(* IEC 61131-3 sources: volt/packages/volt-lsp-iec/test-corpus/pro2193/Device/Plc Logic/Application/09 Misc/Library Manager/L_SUDP_SlaveUpDownloadManager, 64 files *)

(* ---- L_SEMP_ITF_EVENTPARAMETERS.dut ---- *)
TYPE L_SEMP_ITF_EVENTPARAMETERS :
STRUCT
	EVENTPARAMETERS : ARRAY [0..1] OF L_SEMP_ITF_ParameterItem;
END_STRUCT
END_TYPE

(* ---- L_SEMP_ITF_PARAMETERITEM.dut ---- *)
TYPE L_SEMP_ITF_PARAMETERITEM :
STRUCT
	SIZE : BYTE;
	ETYPE : INT;
	VALUE : L_SEMP_ITF_ParaValue;
END_STRUCT
END_TYPE

(* ---- L_SEMP_ITF_PARAVALUE.dut ---- *)
TYPE L_SEMP_ITF_PARAVALUE :
UNION
	DWVALUE : DWORD;
	DNVALUE : DINT;
	FVALUE : REAL;
	STVALUE : STRING;
	DWTEXTLISTID : DWORD;
END_UNION
END_TYPE

(* ---- L_SUDP_BUS_TYPE.dut ---- *)
TYPE L_SUDP_BUS_TYPE :
(
	BUS_CAN := 15,
	BUS_ETC := 64
);
END_TYPE

(* ---- L_SUDP_CONTROL.dut ---- *)
TYPE L_SUDP_CONTROL :
(
	NONE := 0,
	CHECKVERSION := 1,
	DOWNLOAD := 2,
	UPLOAD := 3,
	RESTARTDEVICE := 4,
	PROVIDENEWPARSETCHECKSUM := 5,
	ONLINEPARADOWNLOAD := 6,
	RESTARTDEVICE2 := 7,
	RESTARTDEVICEI750 := 8,
	ABORT := 10
);
END_TYPE

(* ---- L_SUDP_CPAR_FILE_HDR.dut ---- *)
TYPE L_SUDP_CPAR_FILE_HDR :
STRUCT
	DWFILETYPE : DWORD;
	DWVERSION : DWORD;
	DWFILESIZE : DWORD;
	DWVENDOR : DWORD;
	DWPRODUCTTYPE : DWORD;
	DWREVISION : DWORD;
	DWDATAOFF : DWORD;
	DWDATASIZE : DWORD;
	DWFILECRC : DWORD;
END_STRUCT
END_TYPE

(* ---- L_SUDP_ERRORCODES.dut ---- *)
TYPE L_SUDP_ERRORCODES :
(
	NO_ERROR := 0,
	FILE_NOT_FOUND := 1,
	FILE_READ_ERROR := 2,
	PARAM_WRITE_ERROR := 4,
	SLAVE_ERROR := 5,
	PARA_FILE_TYPE_INVALID := 7,
	PARAM_READ_ERROR := 8,
	NO_BUFFER := 9,
	NO_MEMORY := 10,
	WRONG_VERSION_FORMAT := 11,
	ETC_STATE_COULD_NOT_BE_CHANGED := 12,
	GET_FIRMWARE_BINARY_FILE_NAME_FAILED := 13,
	SLAVE_FIRMWARE_UPDATE_FAILED := 14,
	PARAM_SET_UPDATE_FAILED := 15,
	PARAM_SET_FILE_UPLOAD_FAILED := 16,
	PARAM_UPLOAD_FILE_CREATE_FAILED := 17,
	PARAM_WRITE_TO_FILE_FAILED := 18,
	NO_CONFIG_INFORMATION := 19,
	NO_CURRENT_IEC_TASK_INFORMATION := 20,
	NO_FREE_ASYNC_MANAGER := 21,
	FILE_WRITE_ERROR := 22,
	SLAVE_FIRMWARE_UPDATE_HW_INCOMPATIBILITY := 23,
	ERROR_PARAMETERST_UPDATE_FAILED_PARAM_WRITE_ERRORS := 24,
	PARAM_DL_ERROR_FILE_READ_ERROR := 25,
	SLAVE_FW_UPDATE_HW_DIFFERS_NOT_UPDATED := 26
);
END_TYPE

(* ---- L_SUDP_ERRORINDEXSUBINDEX.dut ---- *)
TYPE L_SUDP_ERRORINDEXSUBINDEX :
STRUCT
	WINDEX : WORD;
	WSUBINDEX : BYTE;
END_STRUCT
END_TYPE

(* ---- L_SUDP_MAX_STRING_LENGTH.dut ---- *)
TYPE L_SUDP_MAX_STRING_LENGTH :
(
	FILE_NAME := 50,
	DEVICE_FIRMWARE_VERSION_NUMBER := 30,
	PATH_AND_FILE_NAME := 250,
	FILE_PATH := 200
);
END_TYPE

(* ---- L_SUDP_PAR_DATA_HDR.dut ---- *)
TYPE L_SUDP_PAR_DATA_HDR :
STRUCT
	DWPARTYPE : DWORD;
	DWPARDATAOFF : DWORD;
	DWPARDATSIZE : DWORD;
END_STRUCT
END_TYPE

(* ---- L_SUDP_PAR_FILE_HDR.dut ---- *)
TYPE L_SUDP_PAR_FILE_HDR :
STRUCT
	DWFILETYPE : DWORD;
	DWVERSION : DWORD;
	DWFILESIZE : DWORD;
	DWVENDOR : DWORD;
	DWPRODUCTTYPE : DWORD;
	DWREVISION : DWORD;
	DWDATAOFF : DWORD;
	DWDATASIZE : DWORD;
	DWFILECRC : DWORD;
END_STRUCT
END_TYPE

(* ---- L_SUDP_PAR_FILE_HDR_SEL_PS.dut ---- *)
TYPE L_SUDP_PAR_FILE_HDR_SEL_PS :
STRUCT
	DWFILETYPE : DWORD;
	DWVERSION : DWORD;
	DWFILESIZE : DWORD;
	DWFILECRC : DWORD;
	DWCOUNTPARAMETERSETS : DWORD;
	APARAMETERSETINFO : ARRAY [0..10] OF L_SUDP_PAR_FILE_HDR_SEL_PS_INFO;
END_STRUCT
END_TYPE

(* ---- L_SUDP_PAR_FILE_HDR_SEL_PS_INFO.dut ---- *)
TYPE L_SUDP_PAR_FILE_HDR_SEL_PS_INFO :
STRUCT
	DWPARAMETERSETNUMBER : DWORD;
	DWDATAOFFSET : DWORD;
END_STRUCT
END_TYPE

(* ---- L_SUDP_PARM_ERROR_CODE.dut ---- *)
TYPE L_SUDP_PARM_ERROR_CODE :
STRUCT
	DWERRORCODE : DWORD;
	WINDEX : WORD;
	WSUBINDEX : WORD;
END_STRUCT
END_TYPE

(* ---- L_SUDP_PARM_HDR.dut ---- *)
TYPE L_SUDP_PARM_HDR :
STRUCT
	U16SIZE : UINT;
	U16INDEX : UINT;
	U16SUBINDEX : UINT;
END_STRUCT
END_TYPE

(* ---- L_SUDP_PARM_RECORD.dut ---- *)
TYPE L_SUDP_PARM_RECORD :
STRUCT
	U16SIZE : UINT;
	U16INDEX : UINT;
	U16SUBINDEX : UINT;
	U8DATA : BYTE;
END_STRUCT
END_TYPE

(* ---- L_SUDP_PRM_FILE_READWRITE_STATES.dut ---- *)
TYPE L_SUDP_PRM_FILE_READWRITE_STATES :
(
	NONE,
	WAIT_FILE_SIZE,
	WAIT_READ_FILE_OPEN,
	READ_FILE_HEADERS,
	WRITE_FILE_HEADERS,
	WAIT_WRITE_FILE_OPEN,
	WAIT_READ_PARAM_HEADER,
	WAIT_READ_PARAM_VALUE,
	WAIT_READ_NEXT_PARAM_HEADER_AND_PARAM_VALUE,
	WAIT_WRITE_FILE_PARAMETER,
	WAIT_SET_NEW_FILE_POS_FOR_WRITE_HEADERS,
	WAIT_WRITE_NEW_FILE_HEADERS,
	WAIT_CALC_CHECKSUM,
	WAIT_DELETE_OLD_FILE,
	WAIT_RENAME_NEW_TO_OLD_FILE,
	CLOSE_READ_FILE,
	CLOSE_WRITE_FILE,
	DONE,
	ERROR
);
END_TYPE

(* ---- L_SUDP_STATE.dut ---- *)
TYPE L_SUDP_STATE :
(
	NONE := 0,
	ISREGISTERED := 1,
	DOWNLOADISNECESSARY := 2,
	DOWNLOADISNOTNECESSARY := 3,
	ISBUSY := 4,
	UPDOWNLOADDONE := 5,
	RESTARTDONE := 6,
	NEWCHECKSUMPROVIDED := 7,
	RESTARTDONE2 := 8,
	RESTARTDONEI750 := 9,
	ERROR := 10,
	ABORTED := 20
);
END_TYPE

(* ---- L_SUDP_SUCCESSCODES.dut ---- *)
TYPE L_SUDP_SUCCESSCODES :
(
	SLAVE_FIRMWARE_UPDATE_DONE := 1000,
	SHOW_OLD_FIRMWARE_VERSION := 2000,
	SUDP_DEBUG := 16#2003,
	SUDP_SLAVE_NOT_PRESENT := 16#2004
);
END_TYPE

(* ---- L_SUDP_TRANSFERTYPE.dut ---- *)
TYPE L_SUDP_TRANSFERTYPE :
(
	PARAMETERSETDOWNLOAD := 0,
	PARAMETERSETUPLOAD := 1,
	FIRMWAREDOWNLOAD := 2,
	FIRMWAREDOWNLOAD2 := 3,
	FIRMWAREDOWNLOADI750 := 4
);
END_TYPE

(* ---- DECIMALTOHEXSTRING.pou ---- *)
FUNCTION DECIMALTOHEXSTRING : STRING
VAR_INPUT
	DWVALUE : DWORD;
	NMAXBYTESIZE : INT;
END_VAR
END_FUNCTION

(* ---- GETBOOLEANPROPERTY.pou ---- *)
FUNCTION GETBOOLEANPROPERTY : BOOL
VAR_INPUT
	STKEY : WSTRING;
END_VAR
END_FUNCTION

(* ---- GETCOMPANY.pou ---- *)
FUNCTION GETCOMPANY : WSTRING
END_FUNCTION

(* ---- GETNUMBERPROPERTY.pou ---- *)
FUNCTION GETNUMBERPROPERTY : DINT
VAR_INPUT
	STKEY : WSTRING;
END_VAR
END_FUNCTION

(* ---- GETTEXTPROPERTY.pou ---- *)
FUNCTION GETTEXTPROPERTY : WSTRING
VAR_INPUT
	STKEY : WSTRING;
END_VAR
END_FUNCTION

(* ---- GETTEXTPROPERTY2.pou ---- *)
FUNCTION GETTEXTPROPERTY2 : POINTER TO WSTRING
VAR_INPUT
	STKEY : WSTRING;
END_VAR
END_FUNCTION

(* ---- GETTITLE.pou ---- *)
FUNCTION GETTITLE : WSTRING
END_FUNCTION

(* ---- GETVERSION.pou ---- *)
FUNCTION GETVERSION : VERSION
END_FUNCTION

(* ---- GETVERSIONPROPERTY.pou ---- *)
FUNCTION GETVERSIONPROPERTY : VERSION
VAR_INPUT
	STKEY : WSTRING;
END_VAR
END_FUNCTION

(* ---- L_EXISTALLFILES.pou ---- *)
FUNCTION L_EXISTALLFILES : BOOL
END_FUNCTION

(* ---- L_PATHFIRMWAREFILES.pou ---- *)
FUNCTION L_PATHFIRMWAREFILES : STRING(L_SUDP_MAX_STRING_LENGTH.FILE_PATH)
END_FUNCTION

(* ---- L_PATHPARAMETERSETFILES.pou ---- *)
FUNCTION L_PATHPARAMETERSETFILES : STRING(L_SUDP_MAX_STRING_LENGTH.FILE_PATH)
END_FUNCTION

(* ---- L_SUDP_CRC32FINISH.pou ---- *)
FUNCTION L_SUDP_CRC32FINISH : DWORD
VAR_INPUT
	ULCRC : DWORD;
END_VAR
END_FUNCTION

(* ---- L_SUDP_CRC32INIT.pou ---- *)
FUNCTION L_SUDP_CRC32INIT : DWORD
END_FUNCTION

(* ---- L_SUDP_CRC32UPDATE.pou ---- *)
FUNCTION L_SUDP_CRC32UPDATE : DWORD
VAR_INPUT
	ULCRC : DWORD;
	PDATA : POINTER TO BYTE;
	ULSIZE : __XWORD;
END_VAR
END_FUNCTION

(* ---- L_SUDP_GETBINARYFILENAME.pou ---- *)
FUNCTION L_SUDP_GETBINARYFILENAME : BOOL
VAR_INPUT
	WFIELDBUSMASTERID : WORD;
	WINTERFACE : WORD;
	DNNODEADDRESS : DINT;
	PSBINARYFILENAME : POINTER TO STRING(20);
END_VAR
END_FUNCTION

(* ---- L_SUDP_GETBUFFERINDEX.pou ---- *)
FUNCTION L_SUDP_GETBUFFERINDEX : WORD
VAR_INPUT
	DWLENGTH : DWORD;
	DWTASKINTERVAL : DWORD;
	PERROR : POINTER TO L_SUDP_ErrorCodes;
END_VAR
END_FUNCTION

(* ---- L_SUDP_GETFBCONTROL.pou ---- *)
FUNCTION L_SUDP_GETFBCONTROL : L_SUDP_Control
VAR_INPUT
	HREGISTRATION : CAA.HANDLE;
END_VAR
END_FUNCTION

(* ---- L_SUDP_GETFWDLMODE.pou ---- *)
FUNCTION L_SUDP_GETFWDLMODE : BYTE
END_FUNCTION

(* ---- L_SUDP_GETLEMREGISTRATIONHANDLE.pou ---- *)
FUNCTION L_SUDP_GETLEMREGISTRATIONHANDLE : RTS_IEC_HANDLE
END_FUNCTION

(* ---- L_SUDP_GETPATHBOOTDIRECTORY.pou ---- *)
FUNCTION L_SUDP_GETPATHBOOTDIRECTORY : STRING(L_SUDP_MAX_STRING_LENGTH.FILE_PATH)
END_FUNCTION

(* ---- L_SUDP_GETPATHTEMPDIRECTORY.pou ---- *)
FUNCTION L_SUDP_GETPATHTEMPDIRECTORY : STRING(L_SUDP_MAX_STRING_LENGTH.FILE_PATH)
END_FUNCTION

(* ---- L_SUDP_GETPOINTERTOBUFFER.pou ---- *)
FUNCTION L_SUDP_GETPOINTERTOBUFFER : POINTER TO BYTE
VAR_INPUT
	WBUFFERNUMBER : WORD;
	PERROR : POINTER TO L_SUDP_ErrorCodes;
END_VAR
END_FUNCTION

(* ---- L_SUDP_GETTARGETVERSION.pou ---- *)
FUNCTION L_SUDP_GETTARGETVERSION : BOOL
VAR_INPUT
	ETRANSFERTYPE : L_SUDP_TransferType;
	WFIELDBUSMASTERID : WORD;
	WINTERFACE : WORD;
	DNNODEADDRESS : DINT;
	PSTARGETVERSION : POINTER TO STRING(20);
END_VAR
END_FUNCTION

(* ---- L_SUDP_ISBOOTAPPLICATIONLOADED.pou ---- *)
FUNCTION L_SUDP_ISBOOTAPPLICATIONLOADED : BOOL
END_FUNCTION

(* ---- L_SUDP_REGISTER.pou ---- *)
FUNCTION L_SUDP_REGISTER : CAA.HANDLE
VAR_INPUT
	ETRANSFERTYPE : L_SUDP_TransferType;
	WFIELDBUSMASTERID : WORD;
	WINTERFACE : WORD;
	DNNODEADDRESS : DINT;
END_VAR
END_FUNCTION

(* ---- L_SUDP_RELEASEBUFFERINDEX.pou ---- *)
FUNCTION L_SUDP_RELEASEBUFFERINDEX : BOOL
VAR_INPUT
	WBUFFERINDEX : WORD;
	PERROR : POINTER TO L_SUDP_ErrorCodes;
END_VAR
END_FUNCTION

(* ---- L_SUDP_RELEASEBUFFERINDEXWITHERROR.pou ---- *)
FUNCTION L_SUDP_RELEASEBUFFERINDEXWITHERROR : BOOL
VAR_INPUT
	WBUFFERINDEX : WORD;
	PERROR : POINTER TO L_SUDP_ErrorCodes;
END_VAR
END_FUNCTION

(* ---- L_SUDP_SENDEVENTBUSISPREOP.pou ---- *)
FUNCTION L_SUDP_SENDEVENTBUSISPREOP : BOOL
VAR_INPUT
	WFIELDBUSMASTERID : WORD;
	WINTERFACE : WORD;
END_VAR
END_FUNCTION

(* ---- L_SUDP_SETCANCONFIGURATIONDONE.pou ---- *)
FUNCTION L_SUDP_SETCANCONFIGURATIONDONE : BOOL
VAR_INPUT
	WFIELDBUSMASTERID : WORD;
	WINTERFACE : WORD;
	BYCOUNTOFSLAVE : BYTE;
END_VAR
END_FUNCTION

(* ---- L_SUDP_SETCANISPREOP.pou ---- *)
FUNCTION L_SUDP_SETCANISPREOP
VAR_INPUT
	WFIELDBUSMASTERID : WORD;
	WINTERFACE : WORD;
END_VAR
END_FUNCTION

(* ---- L_SUDP_SETNEWFBERROR.pou ---- *)
FUNCTION L_SUDP_SETNEWFBERROR : BOOL
VAR_INPUT
	HREGISTRATION : CAA.HANDLE;
	EERROR : L_SUDP_ErrorCodes;
END_VAR
END_FUNCTION

(* ---- L_SUDP_SETNEWFBPROGRESS.pou ---- *)
FUNCTION L_SUDP_SETNEWFBPROGRESS : BOOL
VAR_INPUT
	HREGISTRATION : CAA.HANDLE;
	BYPROGRESS : BYTE;
END_VAR
END_FUNCTION

(* ---- L_SUDP_SETNEWFBSTATE.pou ---- *)
FUNCTION L_SUDP_SETNEWFBSTATE : BOOL
VAR_INPUT
	HREGISTRATION : CAA.HANDLE;
	ESTATE : L_SUDP_State;
END_VAR
END_FUNCTION

(* ---- L_SUDP_UPDOWNLOADFBEXIT.pou ---- *)
FUNCTION L_SUDP_UPDOWNLOADFBEXIT : BOOL
VAR_INPUT
	WFIELDBUSMASTERID : WORD;
	WINTERFACE : WORD;
	ETRANSFERTYPE : L_SUDP_TransferType;
END_VAR
END_FUNCTION

(* ---- L_SUDP_UPDOWNLOADFBINIT.pou ---- *)
FUNCTION L_SUDP_UPDOWNLOADFBINIT : BOOL
VAR_INPUT
	WFIELDBUSMASTERID : WORD;
	WINTERFACE : WORD;
	ETRANSFERTYPE : L_SUDP_TransferType;
END_VAR
END_FUNCTION

(* ---- L_SUDP_WRITEERRORMESSAGE.pou ---- *)
FUNCTION L_SUDP_WRITEERRORMESSAGE : BOOL
VAR_INPUT
	HLEMACCESS : RTS_IEC_HANDLE;
	SDEVICENAME : STRING;
	WSLAVEADR : WORD;
	TRANSFERTYPE : L_SUDP_TransferType;
	ERRORCODE : L_SUDP_ErrorCodes;
	PSERRORATTACHMENT : POINTER TO STRING;
END_VAR
END_FUNCTION

(* ---- L_SUDP_WRITEERRORMESSAGEWITHLOGCLASS.pou ---- *)
FUNCTION L_SUDP_WRITEERRORMESSAGEWITHLOGCLASS : BOOL
VAR_INPUT
	HLEMACCESS : RTS_IEC_HANDLE;
	SDEVICENAME : STRING;
	WSLAVEADR : WORD;
	TRANSFERTYPE : L_SUDP_TransferType;
	LOGCLASS : UDINT;
	ERRORCODE : L_SUDP_ErrorCodes;
	PSERRORATTACHMENT : POINTER TO STRING;
END_VAR
END_FUNCTION

(* ---- L_SUDP_WRITELOGMESSAGE.pou ---- *)
FUNCTION L_SUDP_WRITELOGMESSAGE : BOOL
VAR_INPUT
	HLEMACCESS : RTS_IEC_HANDLE;
	SDEVICENAME : STRING;
	WSLAVEADR : WORD;
	TRANSFERTYPE : L_SUDP_TransferType;
	LOGCLASS : UDINT;
	UDILOGID : UDINT;
	PSLOGMESSAGE : POINTER TO STRING;
END_VAR
END_FUNCTION

(* ---- L_SUDP_WRITENEWPARSETCHECKSUM.pou ---- *)
FUNCTION L_SUDP_WRITENEWPARSETCHECKSUM : BOOL
VAR_INPUT
	EBUSTYPE : L_SUDP_BUS_TYPE;
	WNETID : WORD;
	WSLAVEADR : WORD;
	DWFILECRC : DWORD;
END_VAR
END_FUNCTION

(* ---- L_SUDP_WRITESUCCESSMESSAGE.pou ---- *)
FUNCTION L_SUDP_WRITESUCCESSMESSAGE : BOOL
VAR_INPUT
	HLEMACCESS : RTS_IEC_HANDLE;
	SDEVICENAME : STRING;
	WSLAVEADR : WORD;
	TRANSFERTYPE : L_SUDP_TransferType;
	SUCCESSCODE : L_SUDP_SuccessCodes;
	PSATTACHEDTXT : POINTER TO STRING;
END_VAR
END_FUNCTION

(* ---- CALCULATECHECKSUMFROMOPENFILE.pou ---- *)
FUNCTION_BLOCK CALCULATECHECKSUMFROMOPENFILE EXTENDS AsyncBaseClass
VAR_INPUT
	XEXECUTE : BOOL;
	HPARAFILE : RTS_IEC_HANDLE;
	DWFILESIZE : __XWORD;
	PBYBUFFER : POINTER TO BYTE;
	SZBUFFERSIZE : __XWORD;
	DWFILEOFFSETCHECKSUMCALC : DWORD;
	DWPOSITIONCHECKSUM : __XWORD := 32;
END_VAR
VAR_OUTPUT
	XDONE : BOOL;
	XERROR : BOOL;
	EERROR : L_SUDP_ErrorCodes;
	ULCRC32 : UDINT;
END_VAR
VAR
	JOB : RTS_IEC_HANDLE := CAA.gc_hINVALID;
	JOBSTATE : UDINT;
	RESULTTASK : RTS_IEC_RESULT;
	ASYNCJOBPARAM : AsyncJob_Param;
	ASYNCJOBNAME : STRING := 'UploacCalcCRC';
	RESULTASYNCADD : UDINT;
	XEXECUTEOLD : BOOL;
	DWFILEPOS : __XWORD;
	A : INT;
END_VAR
END_FUNCTION_BLOCK

METHOD DOJOB : RTS_IEC_RESULT
END_METHOD

METHOD DUMMYJOB : RTS_IEC_RESULT
END_METHOD

METHOD FB_EXIT : BOOL
VAR_INPUT
	BINCOPYCODE : BOOL;
END_VAR
END_METHOD

METHOD FB_INIT : BOOL
VAR_INPUT
	BINITRETAINS : BOOL;
	BINCOPYCODE : BOOL;
END_VAR
END_METHOD

(* ---- L_SUDP_PRMFILE_READWRITE.pou ---- *)
FUNCTION_BLOCK L_SUDP_PRMFILE_READWRITE
VAR_INPUT
	XEXECUTE : BOOL;
	EBUSTYPE : L_SUDP_BUS_TYPE;
	WNETID : WORD := 0;
	WSLAVEADR : WORD := 1;
	SDEVICENAME : STRING;
	HREGISTRATION : CAA.HANDLE := CAA.gc_hINVALID;
	SFULLFILENAME : STRING(L_SUDP_MAX_STRING_LENGTH.PATH_AND_FILE_NAME);
	UDITIMEOUT : UDINT := 500000;
	DWFILEOFFSETCHECKSUMCALC : DWORD;
END_VAR
VAR_OUTPUT
	XDONE : BOOL;
	XERROR : BOOL;
	EERROR : L_SUDP_ErrorCodes;
	PSATTACHEDERRORTXT : POINTER TO STRING;
END_VAR
VAR
	STATE : L_SUDP_PRM_FILE_READWRITE_STATES := L_SUDP_PRM_FILE_READWRITE_STATES.NONE;
	XEXECUTEOLD : BOOL;
	XREPLACEOLDFILE : BOOL;
	FGETFS : FILE.GetSize;
	FOPEN : FILE.Open;
	FREAD : FILE.Read;
	FWRITE : FILE.Write;
	FCLOSE : FILE.Close;
	FSETPOS : FILE.SetPos;
	FRENAME : FILE.Rename;
	FDELETE : FILE.Delete;
	UDITIMEOUTFILEACCESS : UDINT := 200000;
	CALCCRC : CalculateChecksumFromOpenFile;
	HPARAFILEREAD : CAA.HANDLE;
	HPARAFILEWRITE : RTS_IEC_HANDLE;
	PIOBUFFER : POINTER TO BYTE;
	ADWHEADER : ARRAY [0..((((SIZEOF(L_SUDP_PAR_FILE_HDR) + SIZEOF(L_SUDP_PAR_DATA_HDR)) - 1) / SIZEOF(DWORD)) + 1)] OF DWORD;
	ADWIOBUFFER : ARRAY [0..66] OF DWORD;
	XFIRSTPARAMHEADERWASREAD : BOOL;
	ADWSDOVALUEBUFFER : ARRAY [0..66] OF DWORD;
	DWPARDATASZ : DWORD;
	DWPARDATAPOSITION : DWORD;
	DWNEWPARDATAPOSITION : DWORD;
	PFILEHDR : POINTER TO L_SUDP_PAR_FILE_HDR;
	PPARDATHDR : POINTER TO L_SUDP_PAR_DATA_HDR;
	PARAMHDR : L_SUDP_PARM_HDR;
	PPARAMHDR : POINTER TO L_SUDP_PARM_HDR;
	SZPARAFILESZ : UDINT;
	SDODATALENGTH : UINT;
	SDOVALUEREADDONE : BOOL;
	DWCRC32 : DWORD;
	DWCRC32FILEPOSITION : DWORD;
	MYTESTCOUNTER : INT;
END_VAR
END_FUNCTION_BLOCK

METHOD BEFORESTARTEXECUTION
END_METHOD

METHOD READVALUEFROMFIELDBUS_LOOP : INT
END_METHOD

METHOD READVALUEFROMFIELDBUS_START
VAR_INPUT
	PARAMHDR : POINTER TO L_SUDP_PARM_HDR;
	PBYBUFFER : POINTER TO BYTE;
	SZBUFFERSIZE : UINT;
END_VAR
END_METHOD

METHOD FB_EXIT : BOOL
VAR_INPUT
	BINCOPYCODE : BOOL;
END_VAR
END_METHOD

(* ---- L_SUDP_UPDOWNLOAD.pou ---- *)
FUNCTION_BLOCK L_SUDP_UPDOWNLOAD
VAR_OUTPUT
	ESTATE : L_SUDP_State;
	EERROR : L_SUDP_ErrorCodes;
	BYPROGRESS : BYTE;
END_VAR
VAR
	EBUSTYPE : L_SUDP_BUS_TYPE;
	WNETID : WORD;
	WSLAVEADR : WORD;
	TRANSFERTYPE : L_SUDP_TransferType;
	DWTASKINTERVAL : DWORD;
	PTASKINFO : POINTER TO CmpIecTask.Task_Info2;
	HTASKHANDLE : RTS_IEC_HANDLE;
	ETASKRESULT : RTS_IEC_RESULT;
	BFIRSTINITIALIZEDONE : BOOL;
	BREGISTERTODOWNLOADMANAGERDONE : BOOL;
	HREGISTRATION : CAA.HANDLE := CAA.gc_hINVALID;
	PBYDLUPMGRBUFFER : POINTER TO BYTE;
	WBUFFERINDEX : WORD := SINT_TO_WORD((0 - 1));
	M_HLEMACCESS : RTS_IEC_HANDLE;
	FILE_IO_TIMEOUT_FACTOR : UDINT := 10000;
	ETC_SDO_TIMEOUT_FACTOR : UDINT := 1;
	ETC_FOE_TIMEOUT_FACTOR : UDINT := 5;
	ETC_SET_STATE_TIMEOUT_FACTOR : UDINT := 5;
	PARSET_FILE_TYPE_INVALID : DWORD := 0;
	PARSET_FILE_TYPE_9400 : DWORD := 1;
	PARSET_FILE_TYPE_I700_STORE : DWORD := 2;
	PARSET_FILE_TYPE_I700_ALL : DWORD := 3;
	PARSET_FILE_TYPE_STANDARD : DWORD := 1000;
	INVALID_BUFFER_INDEX : WORD := SINT_TO_WORD((0 - 1));
	LEMACCESSHANDLE : RTS_IEC_HANDLE;
END_VAR
END_FUNCTION_BLOCK

METHOD FB_EXIT : BOOL
VAR_INPUT
	BINCOPYCODE : BOOL;
END_VAR
END_METHOD

METHOD FIRSTINITIALIZE
VAR_INPUT
	PIOCONFIGCONNECTOR : POINTER TO IoConfigConnector;
END_VAR
END_METHOD

METHOD GETPARAMETERSETFILENAME : BOOL
VAR_INPUT
	EFIELDBUSMASTERID : L_SUDP_BUS_TYPE;
	WNETID : WORD;
	WSLAVEADR : WORD;
	PPATHBUFFER : POINTER TO STRING;
END_VAR
VAR_OUTPUT
	BRETC : BOOL := TRUE;
END_VAR
END_METHOD

METHOD GETDWTASKINTERVAL
END_METHOD

METHOD REGISTERFBTODLUPMGR : BOOL
VAR_INPUT
	PIOCONFIGCONNECTOR : POINTER TO IoConfigConnector;
END_VAR
END_METHOD
